(* IEC 61131-3 sources: teller/JD_Teller_LC2_V11/Network/ToolCat, 1 file *)

(* ---- ONE_ToolCat_Table.st ---- *)
#define OBJECTS_CONFIG

FUNCTION GLOBAL TAB ONE_ToolCat
-1$UINT, 0$UINT,
0$UINT, 0$UINT,

14$UDINT,
TO_UDINT(2980745877), "_MyIO", 0$UINT, 3$UINT, 0$UINT,
TO_UDINT(3043040051), "_ScrollArea", 0$UINT, 13$UINT, 0$UINT,
TO_UDINT(1013562163), "_ToolCat", 0$UINT, 2$UINT, 0$UINT,
TO_UDINT(3571405469), "easyFileHandling", 0$UINT, 0$UINT, 1$UINT,
TO_UDINT(3455067800), "easyFileList", 0$UINT, 0$UINT, 0$UINT,
TO_UDINT(2225119864), "MerkerEx", 1$UINT, 18$UINT, 7$UINT,
TO_UDINT(933570811), "RAMex", 1$UINT, 16$UINT, 1$UINT,
TO_UDINT(1850111279), "String", 1$UINT, 10$UINT, 7$UINT,
TO_UDINT(2898603620), "StringInternal", 1$UINT, 70$UINT, 0$UINT,
TO_UDINT(2408581120), "StringRAM", 1$UINT, 10$UINT, 1$UINT,
TO_UDINT(3524110630), "ToolcatHandling", 1$UINT, 1$UINT, 1$UINT,
TO_UDINT(2847896136), "ToolLight", 1$UINT, 1$UINT, 1$UINT,
TO_UDINT(3232495061), "VirtualBaseInit", 1$UINT, 3$UINT, 0$UINT,
TO_UDINT(3928697797), "WisFilter", 0$UINT, 0$UINT, 1$UINT,

1$UINT, TO_UDINT(2590405041), "TOOLLIGHT1\FILEHANDLING",

1$UINT, TO_UDINT(648812873), "TOOLLIGHT1\FILEHANDLING\EXTENSIONFILTER\MERKEREX0",
1$UINT, TO_UDINT(2339572194), "TOOLLIGHT1\FILEHANDLING\FILESTRING\MERKEREX0",
1$UINT, TO_UDINT(3447419793), "TOOLLIGHT1\FILEHANDLING\PATHSTRING\MERKEREX0",
1$UINT, TO_UDINT(2982669661), "TOOLLIGHT1\FILEHANDLING\TOOPENFILESTR\MERKEREX0",
1$UINT, TO_UDINT(1199512598), "TOOLLIGHT1\NEWDIRECTORYSTRING\MERKEREX0",
1$UINT, TO_UDINT(4206854592), "TOOLLIGHT1\NEWFILESTRING\MERKEREX0",
1$UINT, TO_UDINT(928991219), "TOOLLIGHT1\WISFILTER1\STRING2\MERKEREX0",

1$UINT, TO_UDINT(232661701), "TOOLLIGHT1\BOXNAME\DATABUFFER",

1$UINT, TO_UDINT(2537658806), "TOOLLIGHT1\FILEHANDLING\EXTENSIONFILTER",
1$UINT, TO_UDINT(1501854390), "TOOLLIGHT1\FILEHANDLING\FILESTRING",
1$UINT, TO_UDINT(107307615), "TOOLLIGHT1\FILEHANDLING\PATHSTRING",
1$UINT, TO_UDINT(639965759), "TOOLLIGHT1\FILEHANDLING\TOOPENFILESTR",
1$UINT, TO_UDINT(2232942689), "TOOLLIGHT1\NEWDIRECTORYSTRING",
1$UINT, TO_UDINT(738229999), "TOOLLIGHT1\NEWFILESTRING",
1$UINT, TO_UDINT(4005824748), "TOOLLIGHT1\WISFILTER1\STRING2",

1$UINT, TO_UDINT(3536878182), "TOOLLIGHT1\BOXNAME",

1$UINT, TO_UDINT(3362219657), "TOOLLIGHT1\TOOLCATHANDLING",

_NO_ATTR, TO_UDINT(4218591591), "TOOLLIGHT1",

1$UINT, TO_UDINT(2861868813), "TOOLLIGHT1\WISFILTER1",

//Internal connections
0$UDINT,
19$UDINT,
TO_UDINT(0), "PathString", TO_UDINT(11),
TO_UDINT(0), "FileString", TO_UDINT(10),
TO_UDINT(0), "ExtensionFilter", TO_UDINT(9),
TO_UDINT(0), "toOpenFileStr", TO_UDINT(12),
TO_UDINT(9), "MerkerEx0", TO_UDINT(1),
TO_UDINT(10), "MerkerEx0", TO_UDINT(2),
TO_UDINT(11), "MerkerEx0", TO_UDINT(3),
TO_UDINT(12), "MerkerEx0", TO_UDINT(4),
TO_UDINT(13), "MerkerEx0", TO_UDINT(5),
TO_UDINT(14), "MerkerEx0", TO_UDINT(6),
TO_UDINT(15), "MerkerEx0", TO_UDINT(7),
TO_UDINT(16), "DataBuffer", TO_UDINT(8),
TO_UDINT(18), "NewFileString", TO_UDINT(14),
TO_UDINT(18), "ToolcatHandling", TO_UDINT(17),
TO_UDINT(18), "FileHandling", TO_UDINT(0),
TO_UDINT(18), "NewDirectoryString", TO_UDINT(13),
TO_UDINT(18), "WisFilter1", TO_UDINT(19),
TO_UDINT(18), "Boxname", TO_UDINT(16),
TO_UDINT(19), "String2", TO_UDINT(15),
0$UDINT,
23$UDINT,
TO_UDINT(0), "PathString", TO_UDINT(11), "Data",
TO_UDINT(0), "FileString", TO_UDINT(10), "Data",
TO_UDINT(0), "ExtensionFilter", TO_UDINT(9), "Data",
TO_UDINT(0), "toOpenFileString", TO_UDINT(12), "Data",
TO_UDINT(0), "cToolCatLoadInfo", TO_UDINT(17), "LoadInfo",
TO_UDINT(9), "DataBuffer", TO_UDINT(1), "m_udLength",
TO_UDINT(10), "DataBuffer", TO_UDINT(2), "m_udLength",
TO_UDINT(11), "DataBuffer", TO_UDINT(3), "m_udLength",
TO_UDINT(12), "DataBuffer", TO_UDINT(4), "m_udLength",
TO_UDINT(13), "DataBuffer", TO_UDINT(5), "m_udLength",
TO_UDINT(14), "DataBuffer", TO_UDINT(6), "m_udLength",
TO_UDINT(15), "DataBuffer", TO_UDINT(7), "m_udLength",
TO_UDINT(16), "DataBuffer", TO_UDINT(8), "m_udLength",
TO_UDINT(17), "toFileHandling", TO_UDINT(0), "Server0",
TO_UDINT(17), "NewFileString", TO_UDINT(14), "Data",
TO_UDINT(17), "toPathString", TO_UDINT(11), "Data",
TO_UDINT(17), "toFileString", TO_UDINT(10), "Data",
TO_UDINT(17), "toExtensionString", TO_UDINT(9), "Data",
TO_UDINT(17), "toSelFile", TO_UDINT(12), "Data",
TO_UDINT(17), "cFileSelected", TO_UDINT(0), "FileSelectedOK",
TO_UDINT(17), "NewDirectoryString", TO_UDINT(13), "Data",
TO_UDINT(17), "BoxnameOutput", TO_UDINT(16), "Data",
TO_UDINT(19), "ExtFilter", TO_UDINT(9), "Data",

//Initialization values
0$UDINT,
22$UDINT,
TO_UDINT(0), "VerticalLevel", TO_UDINT(1),//|ToolCat.ToolLight1\FileHandling.VerticalLevel;
TO_UDINT(0), "LineWidth", TO_UDINT(0),//|ToolCat.ToolLight1\FileHandling.LineWidth;
TO_UDINT(0), "ExtendedScrollBar", TO_UDINT(1),//|ToolCat.ToolLight1\FileHandling.ExtendedScrollBar;
TO_UDINT(1), "ThreadSafe", TO_UDINT(0),//|ToolCat.ExtensionFilter\FileHandling\ToolLight1\MerkerEx0.ThreadSafe;
TO_UDINT(2), "ThreadSafe", TO_UDINT(0),//|ToolCat.FileString\FileHandling\ToolLight1\MerkerEx0.ThreadSafe;
TO_UDINT(3), "ThreadSafe", TO_UDINT(0),//|ToolCat.PathString\FileHandling\ToolLight1\MerkerEx0.ThreadSafe;
TO_UDINT(4), "ThreadSafe", TO_UDINT(0),//|ToolCat.toOpenFileStr\FileHandling\ToolLight1\MerkerEx0.ThreadSafe;
TO_UDINT(5), "ThreadSafe", TO_UDINT(0),//|ToolCat.NewDirectoryString\ToolLight1\MerkerEx0.ThreadSafe;
TO_UDINT(6), "ThreadSafe", TO_UDINT(0),//|ToolCat.NewFileString\ToolLight1\MerkerEx0.ThreadSafe;
TO_UDINT(7), "ThreadSafe", TO_UDINT(0),//|ToolCat.String2\WisFilter1\ToolLight1\MerkerEx0.ThreadSafe;
TO_UDINT(8), "ThreadSafe", TO_UDINT(0),//|ToolCat.Boxname\ToolLight1\DataBuffer.ThreadSafe;
TO_UDINT(9), "SingleRealloc", TO_UDINT(1),//|ToolCat.FileHandling\ToolLight1\ExtensionFilter.SingleRealloc;
TO_UDINT(10), "SingleRealloc", TO_UDINT(1),//|ToolCat.FileHandling\ToolLight1\FileString.SingleRealloc;
TO_UDINT(11), "SingleRealloc", TO_UDINT(1),//|ToolCat.FileHandling\ToolLight1\PathString.SingleRealloc;
TO_UDINT(12), "SingleRealloc", TO_UDINT(1),//|ToolCat.FileHandling\ToolLight1\toOpenFileStr.SingleRealloc;
TO_UDINT(13), "SingleRealloc", TO_UDINT(1),//|ToolCat.ToolLight1\NewDirectoryString.SingleRealloc;
TO_UDINT(14), "SingleRealloc", TO_UDINT(1),//|ToolCat.ToolLight1\NewFileString.SingleRealloc;
TO_UDINT(15), "SingleRealloc", TO_UDINT(1),//|ToolCat.WisFilter1\ToolLight1\String2.SingleRealloc;
TO_UDINT(16), "SingleRealloc", TO_UDINT(1),//|ToolCat.ToolLight1\Boxname.SingleRealloc;
TO_UDINT(17), "Filter", TO_UDINT(1),//|ToolCat.ToolLight1\ToolcatHandling.Filter;
TO_UDINT(17), "cWindowNrFileExists", TO_UDINT(106),//|ToolCat.ToolLight1\ToolcatHandling.cWindowNrFileExists;
TO_UDINT(18), "cWindowNrFileExists", TO_UDINT(106),//|ToolCat.ToolLight1.cWindowNrFileExists;

//Symbolic initialization values
0$UDINT,
0$UDINT,

//Initialization of string values
0$UDINT,
1$UDINT,
TO_UDINT(11), "", 0$UINT, TO_UINT(OFF(L1)-OFF(L0)), L0:"C:\REC\BOXES\",L1://|ToolCat.FileHandling\ToolLight1\PathString.Data;

//Configuration of tasks (RealTime, Cyclic, Background)
0$UDINT,
0$UDINT,

0$UDINT,
0$UDINT,

0$UDINT,
1$UDINT,
TO_UDINT(17), (100)$UDINT, 4194305$DINT, 	//TOOLLIGHT1\TOOLCATHANDLING

//External connections
0$UDINT,
2$UDINT,
TO_UDINT(18), "Lse", C_DIR, TO_UDINT(299963966), "Lse","Lse",
TO_UDINT(18), "Lse0", C_DIR, TO_UDINT(299963966), "Lse","Lse",

//Magic internal connections
0$UDINT,
3$UDINT,
TO_UDINT(0), "Lse", TO_UDINT(18), "Lse0",
TO_UDINT(8), "UseFile", TO_UDINT(16), "UseFile",
TO_UDINT(17), "cWindowNrFileExists", TO_UDINT(18), "cWindowNrFileExists",

//Configuration of timeslots of tasks (RealTime, Cyclic)
#ifdef __LSLLDR_TIMESLOTS__
0$UDINT,
0$UDINT,

0$UDINT,
0$UDINT,

#endif //__LSLLDR_TIMESLOTS__

//MultiMaster connections
#ifdef __LSLLDR_MULTIMASTER__
0$UDINT,
0$UDINT,
#endif //__LSLLDR_MULTIMASTER__

END_FUNCTION
